TEXTLIST TextList_E_Line_Source
  0 = 'Drain'
  1 = 'Tank_A'
  2 = 'Tank_B'
  3 = 'TapWater'
  4 = 'FillWater'
  5 = 'CIP'
   = ''
END_TEXTLIST

(* stored: Version 1.1.0.1, ProductVersion 3.1.4024.12
   TextList TextList_E_Line_Source: Id {4ebd7c6c-3e1a-475b-a824-4802b7d66b7f} *)
